Fanuc KAREL source: KT00685.KL

PROGRAM KT00685
%NOLOCKGROUP
VAR
  P1: JOINTPOS
  P2: JOINTPOS
  OUT: INTEGER
BEGIN
  OUT = - P1
END KT00685
